(* IEC 61131-3 sources: codesys-to-s7/tests/corpus/C2S7-GFX-GOTO/neg, 1 file *)

(* ---- input.st ---- *)
FUNCTION_BLOCK FB_J
VAR_INPUT
    a : BOOL;
END_VAR
VAR
    i : INT;
END_VAR
IF NOT a THEN
    i := 1;
END_IF
i := i + 2;
END_FUNCTION_BLOCK
